// TIA Portal V20 export
FUNCTION "AchsePOS_BIT" : Void   // FC109, STL
TITLE = Achsenposition IST-POS mit Vorgabe vergleichen und Bit setzen
{ S7_Optimized_Access := 'FALSE' }
// stored: AutoNumber false
   VAR_INPUT
      ISTPOS_Achse : Real;   // Istposition der Achse
      POS_Vorgabe : Real;   // Achsposition die als Bit-Position benötigt wird
      Max_Abweichung : Real;   // +/- Abweichung in mm zur Achsposition
   END_VAR
   VAR_OUTPUT
      POS_OK : Bool;   // Wenn Istposition im Fenster POS_Vorgabe +/- MAX Abweichung ist dann VKE=1
   END_VAR
BEGIN

NETWORK
TITLE = Wenn Istposition im Fenster POS_Vorgabe +/- MAX Abweichung ist dann VKE=1
      A(;
      L     #ISTPOS_Achse;
      L     #POS_Vorgabe;
      -R;
      ABS;
      L     #Max_Abweichung;
      <=R;
      );
      =     #POS_OK;
END_FUNCTION
